(* CODESYS project Speed.xml

Project tree, tasks and I/O mapping:
*)

// Speed
PROPERTY Speed : INT
END_PROPERTY
